(* Logix 5000 project; controller TFF vendor 1 type 14 code 107 rev 34.11; software revision 34.03; part 14 of 36 *)
(* tags used below, declared in another part *)
   ActionCode : DINT;   // Action Code
   ActionValue : REAL;   // Action Value
   Boolean : DINT;   // Boolean Operator
   Branch : BOOL;   // Conditional Branch Flag
   Clear : BOOL;   // Clear Operation Table Flag
   Criteria1BoolValue : BOOL;   // Criteria 1 Discrete Value
   Criteria1Code : DINT;   // Criteria 1 Code
   Criteria1Met : BOOL;   // Criteria 1 Met
   Criteria1Operator : DINT;   // Criteria 1 Operator
   Criteria1RealValue : REAL;   // Criteria 1 Real Value
   Criteria1Type : BOOL;   // Criteria 1 Type 0=Real, 1=Boolean
   Criteria1Value : REAL;   // Criteria 1 Value
   Criteria2BoolValue : BOOL;   // Criteria 2 Discrete Value
   Criteria2Code : DINT;   // Criteria 2 Code
   Criteria2Met : BOOL;   // Criteria 2 Met
   Criteria2Operator : DINT;   // Criteria 2 Operator
   Criteria2RealValue : REAL;   // Criteria 2 Real Value
   Criteria2Type : BOOL;   // Criteria 2 Type 0=Real, 1=Boolean
   Criteria2Value : REAL;   // Criteria 2 Value
   CriteriaMet : BOOL;   // Criteria Met
   DateTime : DINT[7];   // Date and Time
   ErrorCheck : BOOL;   // Error Check Flag
   LastStep : DINT;   // Last Step
   NextStep : DINT;   // Next Step
   PendingStep : DINT;   // Current Step
   PhaseNumber : DINT;   // Phase FOR NEXT Index
   Run : BOOL;   // Operation Run Status
   sColon : STRING4;   // Colon separator String
   sComma : STRING4;   // Comma String
   sDateTime : STRING25;   // Date and Time String
   sPeriod : STRING4;   // Timer separator String
   sTemp : STRING50;   // Temp String
   Structure : DINT;   // Structure code
   sZero : STRING4;   // Zero String
   Tag : DINT;   // Tag value
   Tenths : DINT;   // Thents (Date and Time management)
   ThisStep : DINT;   // This Step (Error management)
   Value : REAL;   // Temp Value
   AlarmControl : AlarmControl;   // Alarm Control
   CCPSystem : CCPSystem;   // CCP System Data
   CPU_Scanning : BOOL;   // System Scanning Flag
   FirstScanComplete : BOOL;   // First Scan Complete Flag
   HoldTime : ALIAS FOR Timers[20];   // Hold Time
   Operation : Operation[6,251];   // Operation Table
   Phase : Phases[6];   // Phase Control Array
   Phase0 : ALIAS FOR Phase[0];   // Phase 0
   Phase0_Totalizer_Feed : ALIAS FOR PhaseTotalizer[0];   // Phase 0 Total Feed
   Phase0_Totalizer_Filtrate : ALIAS FOR PhaseTotalizer[6];   // Phase 0 Total Filtrate
   Phase0_Totalizer_Retentate : ALIAS FOR PhaseTotalizer[12];   // Phase 0 Total Retentate
   PhaseTotalizer : PhaseTotalizer[18];   // Phase Totalizers Array
   PLCFault : FaultRecordType;   // PLC Major Fault Record
   ProcedureTime : ALIAS FOR Timers[19];   // Procedure Time
   Prompt : Prompt[7];   // Prompt Array
   TimerControl : TimerControl;   // Timer Control
   Timers : Timers[22];   // Timer Array
   Totalizer : Totalizers[20];   // Totalizers Array
   YA10 : ALIAS FOR DigitalPoint[59];   // PLC Program Major Fault
(* CCPSystem, continued *)

ROUTINE DateTime   (* structured text *)
// System Date and Time Routine
   (* =======================================================================
   	DateTime : 	This routine returns a string value of date and time in the format "MMDDYYYY,HH:MM:SS.x,".
   				The result is stored in the program tag sDateTime.
   				This string will be used by the BufferEvents and BufferSteps routines for time stamping.
   
   	List of treatments
   		- Get system date and time with GSV instruction
   		- Convert the date and time in DINT format to string format
   
   -----------------------------------------------------------------------------------------------------------------------------------------------------
   	History
   		2019-AUG-13 - ACTEMIUM - B. Roch - Initial version for Candidate Release 3.00.00.00.a
   =========================================================================*)
   
   
   (* Get system date and time with GSV instruction
   =========================================================================*)
   
   (*Get the current date and time from the processor*)
   (*The date and time are stored in an array of 7 values*)
   	GSV (WALLCLOCKTIME, , DateTime, DateTime[0]);
   
   (* Convert the date and time in DINT format to string format
   =========================================================================*)
   (*Month*)
   	DTOS (DateTime[1], sDateTime);
   	(*Add leading zero if value is 1 character*)
   	IF sDateTime.LEN = 1 Then;
   		CONCAT (sZero, sDateTime, sDateTime);
   	END_IF;
   (*Day*)
   	DTOS (DateTime[2], sTemp);
   	(*Add leading zero if value is 1 character*)
   	IF sTemp.LEN = 1 Then;
   		CONCAT (sZero, sTemp, sTemp);
   	END_IF;
   	CONCAT (sDateTime, sTemp, sDateTime);
   (*Year*)
   	DTOS (DateTime[0], sTemp);
   	CONCAT (sDateTime, sTemp, sDateTime);
   	CONCAT (sDateTime, sComma, sDateTime);
   (*Hours*)
   	DTOS (DateTime[3], sTemp);
   	(*Add leading zero if value is 1 character*)
   	IF sTemp.LEN = 1 Then;
   		CONCAT (sZero, sTemp, sTemp);
   	END_IF;
   	CONCAT (sDateTime, sTemp, sDateTime);
   	CONCAT (sDateTime, sColon, sDateTime);
   (*Minutes*)
   	DTOS (DateTime[4], sTemp);
   	(*Add leading zero if value is 1 character*)
   	IF sTemp.LEN = 1 Then;
   		CONCAT (sZero, sTemp, sTemp);
   	END_IF;
   	CONCAT (sDateTime, sTemp, sDateTime);
   	CONCAT (sDateTime, sColon, sDateTime);
   (*Seconds*)
   	DTOS (DateTime[5], sTemp);
   	(*Add leading zero if value is 1 character*)
   	IF sTemp.LEN = 1 Then;
   		CONCAT (sZero, sTemp, sTemp);
   	END_IF;
   	CONCAT (sDateTime, sTemp, sDateTime);
   	CONCAT (sDateTime, sPeriod, sDateTime);
   (*Tenth Seconds*)
   	(*Round the microseconds value to tenths seconds*)
   	Tenths := DateTime[6] / 100000;
   	DTOS (Tenths, sTemp);
   	CONCAT (sDateTime, sTemp, sDateTime);
   	CONCAT (sDateTime, sComma, sDateTime);
   
END_ROUTINE

ROUTINE Error   (* structured text *)
// Step Error Checking
   (* =======================================================================
   	Error : This routine loops through all steps of one phase per processor scan to detect an error
   
   	List of treatments
   		- Initialize
   		- Error check processing
   		- Error found
   		- No error found
   
   -----------------------------------------------------------------------------------------------------------------------------------------------------
   	History
   		2019-AUG-13 - ACTEMIUM - B. Roch - Initial version for Candidate Release 3.00.00.00.a
   		2019-SEP-09 - ACTEMIUM - Q. Spindler - Modifications for Candidate Release 3.00.00.00.c
   					- Change Error check for Criterias and Action Value to -999999.99
   =========================================================================*)
   
   
   (* Initialize
   =========================================================================*)
   (*Initialize error check values first time*)
   IF NOT ErrorCheck THEN;
   	CCPSystem.Error := 0;
   	CCPSystem.ErrorStep:= 0;
   	CCPSystem.ErrorPhase := 0;
   	PhaseNumber := 0;
   	ErrorCheck := 1;
   ELSE;
   	PhaseNumber := PhaseNumber + 1;
   END_IF;
   (* PhaseNumber := 5;*)
   (*Reset the total and last step values*)
   Phase[PhaseNumber].TotalSteps := 0;
   LastStep := 0;
   
   (* Error check processing
   =========================================================================*)
   (*Loop through the steps.  If step number is zero, complete*)
   FOR PendingStep := 1 TO 250 DO;
   	IF Operation[PhaseNumber, PendingStep].Step = 0 THEN;
   		EXIT;
   	END_IF;
   
   	(*Step Number Error Check*)
   	(*Verify step number is equal to or one greater than the previous step number*)
   	ThisStep := Operation[PhaseNumber, PendingStep].Step;
   	IF ThisStep <> LastStep + 1 AND ThisStep <> LastStep THEN;
   		CCPSystem.Error := 1;
   		EXIT;
   	END_IF;
   	LastStep := ThisStep;
   	Phase[PhaseNumber].TotalSteps := PendingStep;
   
   	(*Criteria 1 Error Check*)
   	JSR (Criteria1);
   	IF CCPSystem.Error <> 0 THEN;
   		EXIT;
   	END_IF;
   	IF Criteria1Operator <> 0 AND Criteria1Operator <> 1 AND Criteria1Operator <> 2 AND Criteria1Operator <> 4 THEN;
   		CCPSystem.Error := 3;
   		EXIT;
   	ELSIF Boolean > 2 THEN;
   		CCPSystem.Error := 4;
   		EXIT;
   	ELSIF Criteria1Value = -999999.99 THEN;
   		CCPSystem.Error := 9;
   		EXIT;
   	END_IF;
   
   	(*Criteria 2 Error Check*)
   	JSR (Criteria2);
   	IF CCPSystem.Error <> 0 THEN;
   		EXIT;
   	END_IF;
   	IF Criteria2Operator <> 0 AND Criteria2Operator <> 1 AND Criteria2Operator <> 2 AND Criteria2Operator <> 4 THEN;
   		CCPSystem.Error := 6;
   		EXIT;
   	ELSIF Criteria2Value = -999999.99 THEN;
   		CCPSystem.Error := 10;
   		EXIT;
   	END_IF;
   
   	(*Action Error Check*)
   	JSR (Action);
   	IF CCPSystem.Error <> 0 THEN;
   		EXIT;
   	END_IF;
   	IF ActionValue = -999999.99 THEN;
   		CCPSystem.Error := 11;
   		EXIT;
   	END_IF;
   
   	(*Label Error Check*)
   	IF  Operation[PhaseNumber, PendingStep].Label > 20 THEN;
   		CCPSystem.Error := 8;
   		EXIT;
   	END_IF;
   END_FOR;
   
   (* Error found
   =========================================================================*)
   (*Error Found. Set state to 13, record step and phase number, clear error check flag*)
   IF CCPSystem.Error <> 0 THEN;
   	ErrorCheck := 0;
   	CCPSystem.State := 13;
   	CCPSystem.ErrorStep := PendingStep;
   	CCPSystem.ErrorPhase := PhaseNumber;
   END_IF;
   
   (* No error found
   =========================================================================*)
   (*Complete with no errors. Set state to 0 and clear error check flag*)
   IF PhaseNumber = 5 AND CCPSystem.Error = 0 THEN;
   	ErrorCheck := 0;
   	CCPSystem.State := 0;
   	DTOS (0, CCPSystem.BufferSteps[0]);
   END_IF;
END_ROUTINE

ROUTINE FaultRoutine   (* ladder *)
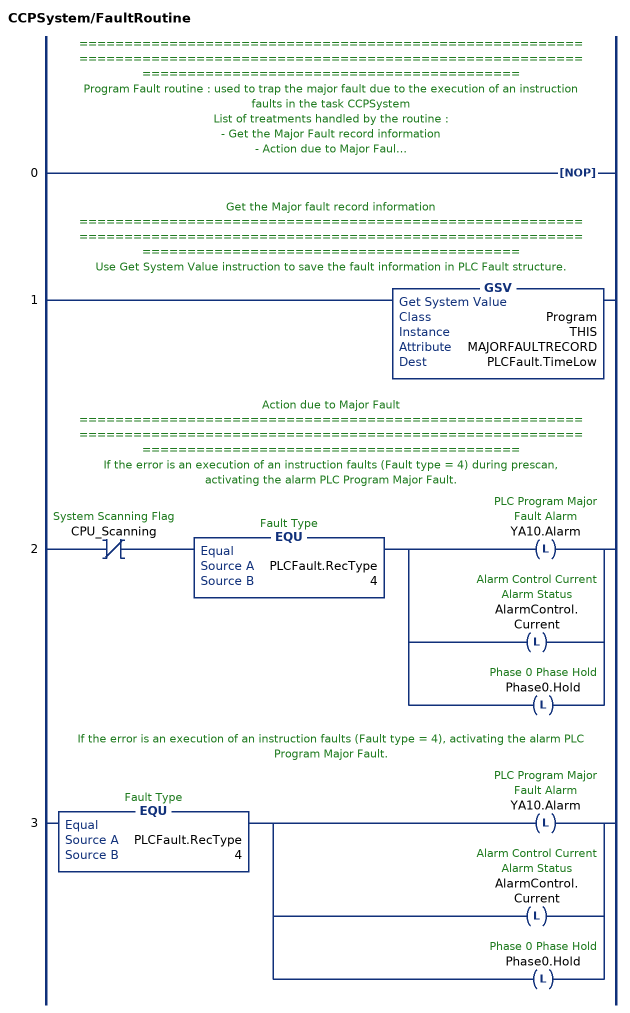
   // ==========================================================================================================================================================
   //                                                            Program Fault routine : used to trap the major fault due to the execution of an instruction faults in the task CCPSystem
   //                                                     List of treatments handled by the routine :
   //                                                          - Get the Major Fault record information
   //                                                          - Action due to Major Fault
   //                                                     -----------------------------------------------------------------------------------------------------------------------------------------------------
   //                                                     History
   //                                                         2019-AUG-13 - Actemium - B. Roch - Initial version for Candidate Release 3.00.00.00.a
   // ==========================================================================================================================================================
   0: NOP();
   // Get the Major fault record information
   // ==========================================================================================================================================================
   // Use Get System Value instruction to save the fault information in PLC Fault structure.
   1: GSV(Program,THIS,MAJORFAULTRECORD,PLCFault.TimeLow);
   // Action due to Major Fault
   // ==========================================================================================================================================================
   // If the error is an execution of an instruction faults (Fault type = 4) during prescan, activating the alarm PLC Program Major Fault.
   2: XIO(CPU_Scanning)EQU(PLCFault.RecType,4)[OTL(YA10.Alarm) ,OTL(AlarmControl.Current) ,OTL(Phase0.Hold) ];
   // If the error is an execution of an instruction faults (Fault type = 4), activating the alarm PLC Program Major Fault.
   3: EQU(PLCFault.RecType,4)[OTL(YA10.Alarm) ,OTL(AlarmControl.Current) ,OTL(Phase0.Hold) ];
END_ROUTINE

ROUTINE MainRoutine   (* ladder *)
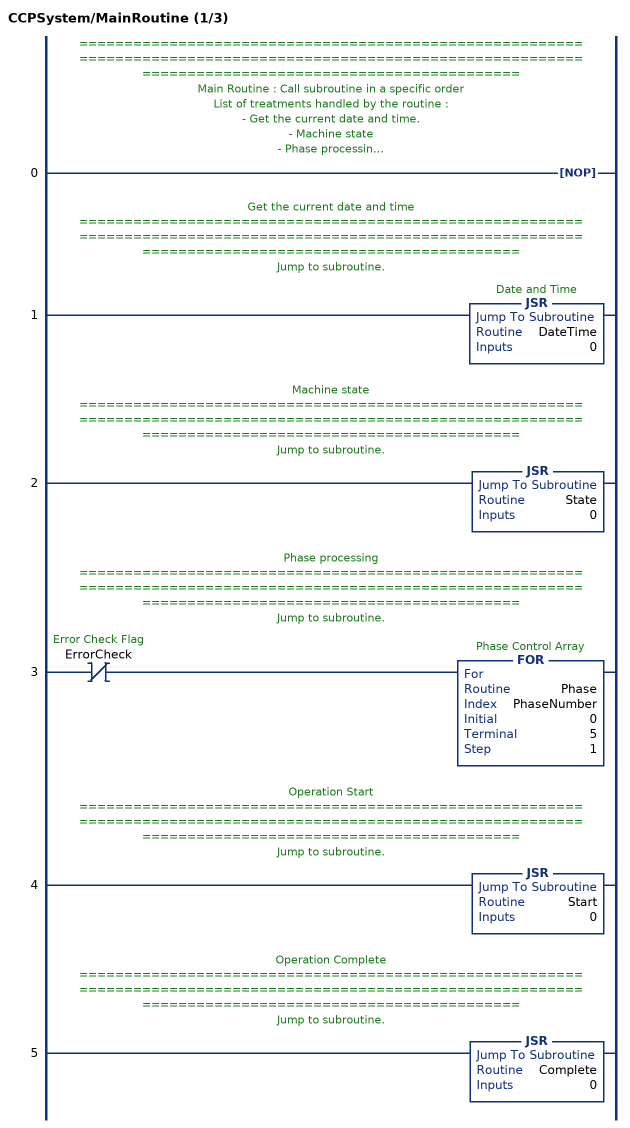
   // ==========================================================================================================================================================
   //                                                                                                            Main Routine : Call subroutine in a specific order
   //                                                     List of treatments handled by the routine :
   //                                                          - Get the current date and time.
   //                                                          - Machine state
   //                                                          - Phase processing
   //                                                          - Operation Start
   //                                                          - Operation Complete
   //                                                          - Procedure timer and totalizer - Hold timer
   //                                                          - Event Log
   //                                                          - CCP System watchdog
   //                                                     -----------------------------------------------------------------------------------------------------------------------------------------------------
   //                                                     History
   //                                                          2019-AUG-13 - Actemium - B. Roch - Initial version for Candidate Release 3.00.00.00.a
   // 2020-SEP-30 - Merck - Q.Spindler - Modifications for Candidate Release 3.00.00.01.a
   // - Add Retentate totalizer
   // ========================================================================================================================================================
   0: NOP();
   // Get the current date and time
   // ==========================================================================================================================================================
   // Jump to subroutine.
   1: JSR(DateTime,0);
   // Machine state
   // ==========================================================================================================================================================
   // Jump to subroutine.
   2: JSR(State,0);
   // Phase processing
   // ==========================================================================================================================================================
   // Jump to subroutine.
   3: XIO(ErrorCheck)FOR(Phase,PhaseNumber,0,5,1);
   // Operation Start
   // ==========================================================================================================================================================
   // Jump to subroutine.
   4: JSR(Start,0);
   // Operation Complete
   // ==========================================================================================================================================================
   // Jump to subroutine.
   5: JSR(Complete,0);
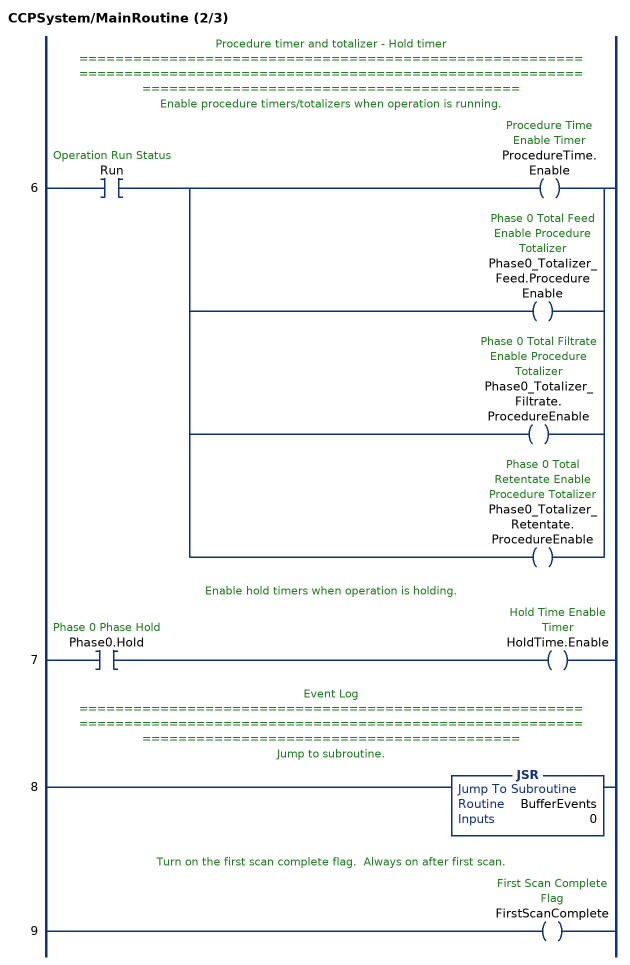
   // Procedure timer and totalizer - Hold timer
   // ==========================================================================================================================================================
   // Enable procedure timers/totalizers when operation is running.
   6: XIC(Run)[OTE(ProcedureTime.Enable) ,OTE(Phase0_Totalizer_Feed.ProcedureEnable) ,OTE(Phase0_Totalizer_Filtrate.ProcedureEnable) ,OTE(Phase0_Totalizer_Retentate.ProcedureEnable) ];
   // Enable hold timers when operation is holding.
   7: XIC(Phase0.Hold)OTE(HoldTime.Enable);
   // Event Log
   // ==========================================================================================================================================================
   // Jump to subroutine.
   8: JSR(BufferEvents,0);
   // Turn on the first scan complete flag.  Always on after first scan.
   9: OTE(FirstScanComplete);
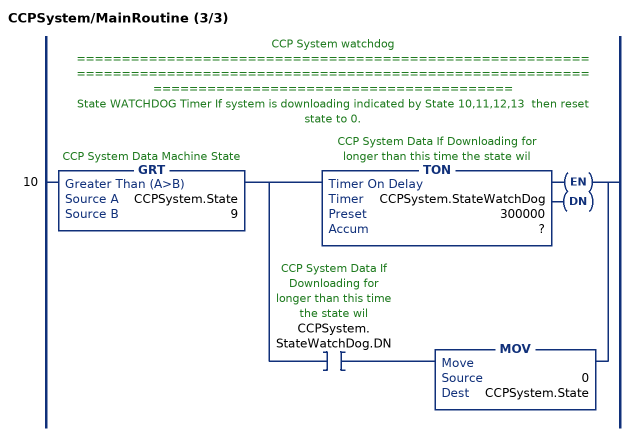
   // CCP System watchdog
   // ==========================================================================================================================================================
   // State WATCHDOG Timer If system is downloading indicated by State 10,11,12,13  then reset state to 0.
   10: GRT(CCPSystem.State,9)[TON(CCPSystem.StateWatchDog,?,?) ,XIC(CCPSystem.StateWatchDog.DN) MOV(0,CCPSystem.State) ];
END_ROUTINE

ROUTINE Phase   (* ladder *)
// Phase Processing Routine
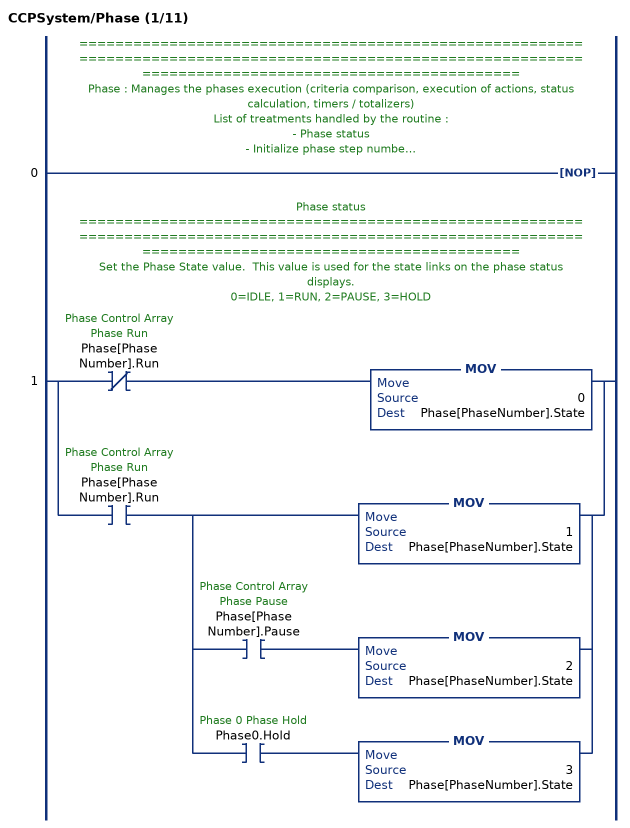
   // ==========================================================================================================================================================
   //                                                                   Phase : Manages the phases execution (criteria comparison, execution of actions, status calculation, timers / totalizers)
   //                                                     List of treatments handled by the routine :
   //                                                          - Phase status
   //                                                          - Initialize phase step number
   //                                                          - Phase Timer / Toalizer
   //                                                          - Phase Stop
   //                                                          - Criteria 1 processing
   //                                                          - Criteria 2 processing
   //                                                          - Jump Step
   //                                                          - Criteria met
   //                                                          - Phase Pause
   //                                                          - Prompt processing
   //                                                          - Branch step processing
   //                                                          - Action processing
   //                                                          - Update step number
   //                                                          - Reset step timer and totalizer
   //                                                     -----------------------------------------------------------------------------------------------------------------------------------------------------
   //                                                     History
   //                                 2019-AUG-13 - Actemium - B. Roch - Initial version for Candidate Release 3.00.00.00.a
   //                                2020-SEP-14 - Merck - Q. Spindler - Modifications for Candidate Release 3.00.00.01.a
   //                                                      - Replace TimerControl.Tick by TimerControl.TickMainTask
   // - Add Retentate totalizer
   // 		               2021-MAY-03 - DAVIDSON- Ch. ARBOGAST - Modifications for Candidate Release 3.01.00.00.a
   //  			- on rung 19 "Reset the step timers...", add "CLR Phase[PhaseNumber].Crit1MetTime"
   //                                          2023-FEB-07 - Davidson - Ch.ARBOGAST - Modifications for Candidate Release 3.02.00.00.a
   //                                                                       - Rung 8. add Hold condition for criteria 1 met Timer (block timer if system in Hold)
   // ========================================================================================================================================================
   0: NOP();
   // Phase status
   // ==========================================================================================================================================================
   // Set the Phase State value.  This value is used for the state links on the phase status displays.
   // 0=IDLE, 1=RUN, 2=PAUSE, 3=HOLD
   1: [XIO(Phase[PhaseNumber].Run) MOV(0,Phase[PhaseNumber].State) ,XIC(Phase[PhaseNumber].Run) [MOV(1,Phase[PhaseNumber].State) ,XIC(Phase[PhaseNumber].Pause) MOV(2,Phase[PhaseNumber].State) ,XIC(Phase0.Hold) MOV(3,Phase[PhaseNumber].State) ] ];
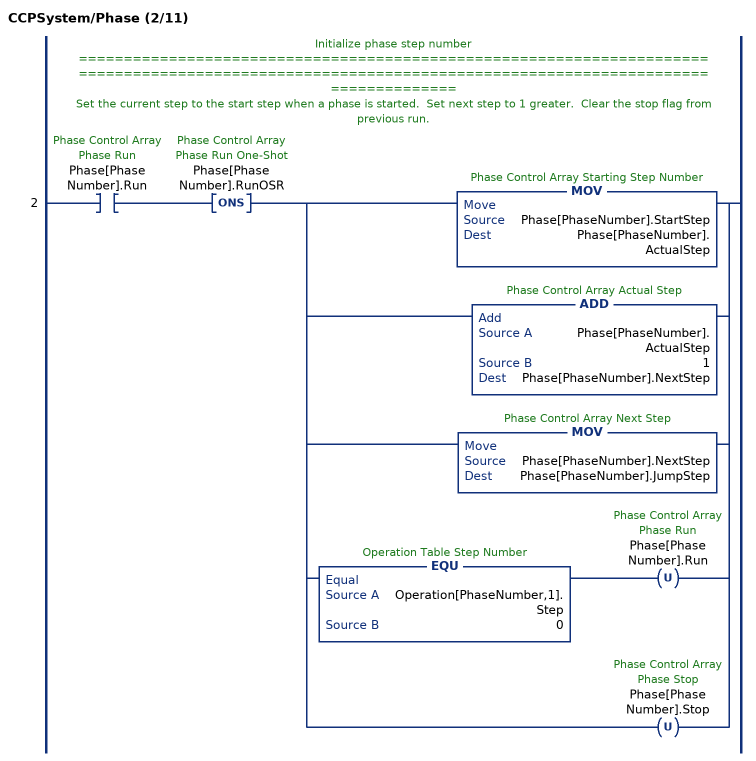
   // Initialize phase step number
   // ==========================================================================================================================================================
   // Set the current step to the start step when a phase is started.  Set next step to 1 greater.  Clear the stop flag from previous run.
   2: XIC(Phase[PhaseNumber].Run)ONS(Phase[PhaseNumber].RunOSR)[MOV(Phase[PhaseNumber].StartStep,Phase[PhaseNumber].ActualStep) ,ADD(Phase[PhaseNumber].ActualStep,1,Phase[PhaseNumber].NextStep) ,MOV(Phase[PhaseNumber].NextStep,Phase[PhaseNumber].JumpStep) ,EQU(Operation[PhaseNumber,1].Step,0) OTU(Phase[PhaseNumber].Run) ,OTU(Phase[PhaseNumber].Stop) ];
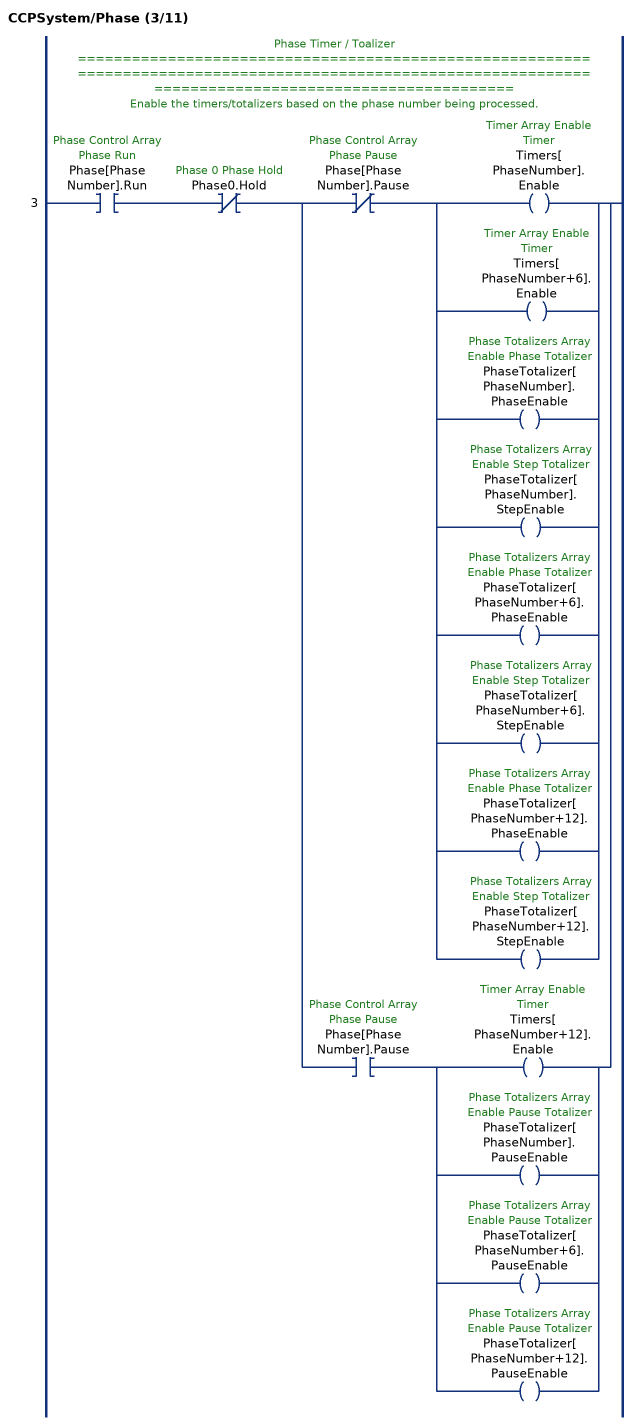
   // Phase Timer / Toalizer
   // ==========================================================================================================================================================
   // Enable the timers/totalizers based on the phase number being processed.
   3: XIC(Phase[PhaseNumber].Run)XIO(Phase0.Hold)[XIO(Phase[PhaseNumber].Pause) [OTE(Timers[PhaseNumber].Enable) ,OTE(Timers[PhaseNumber+6].Enable) ,OTE(PhaseTotalizer[PhaseNumber].PhaseEnable) ,OTE(PhaseTotalizer[PhaseNumber].StepEnable) ,OTE(PhaseTotalizer[PhaseNumber+6].PhaseEnable) ,OTE(PhaseTotalizer[PhaseNumber+6].StepEnable) ,OTE(PhaseTotalizer[PhaseNumber+12].PhaseEnable) ,OTE(PhaseTotalizer[PhaseNumber+12].StepEnable) ] ,XIC(Phase[PhaseNumber].Pause) [OTE(Timers[PhaseNumber+12].Enable) ,OTE(PhaseTotalizer[PhaseNumber].PauseEnable) ,OTE(PhaseTotalizer[PhaseNumber+6].PauseEnable) ,OTE(PhaseTotalizer[PhaseNumber+12].PauseEnable) ] ];
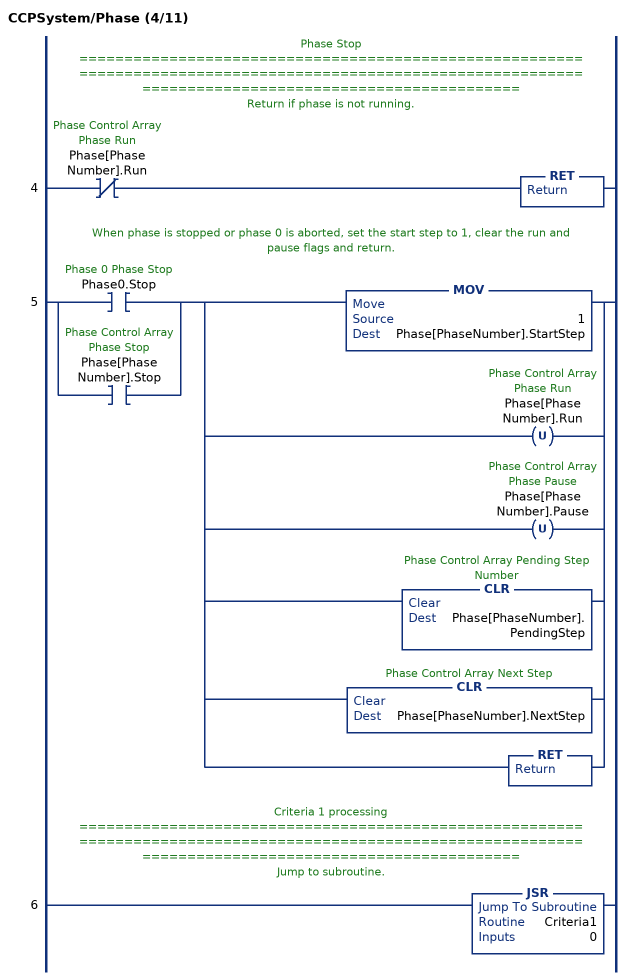
   // Phase Stop
   // ==========================================================================================================================================================
   // Return if phase is not running.
   4: XIO(Phase[PhaseNumber].Run)RET();
   // When phase is stopped or phase 0 is aborted, set the start step to 1, clear the run and pause flags and return.
   5: [XIC(Phase0.Stop) ,XIC(Phase[PhaseNumber].Stop) ][MOV(1,Phase[PhaseNumber].StartStep) ,OTU(Phase[PhaseNumber].Run) ,OTU(Phase[PhaseNumber].Pause) ,CLR(Phase[PhaseNumber].PendingStep) ,CLR(Phase[PhaseNumber].NextStep) ,RET() ];
   // Criteria 1 processing
   // ==========================================================================================================================================================
   // Jump to subroutine.
   6: JSR(Criteria1,0);
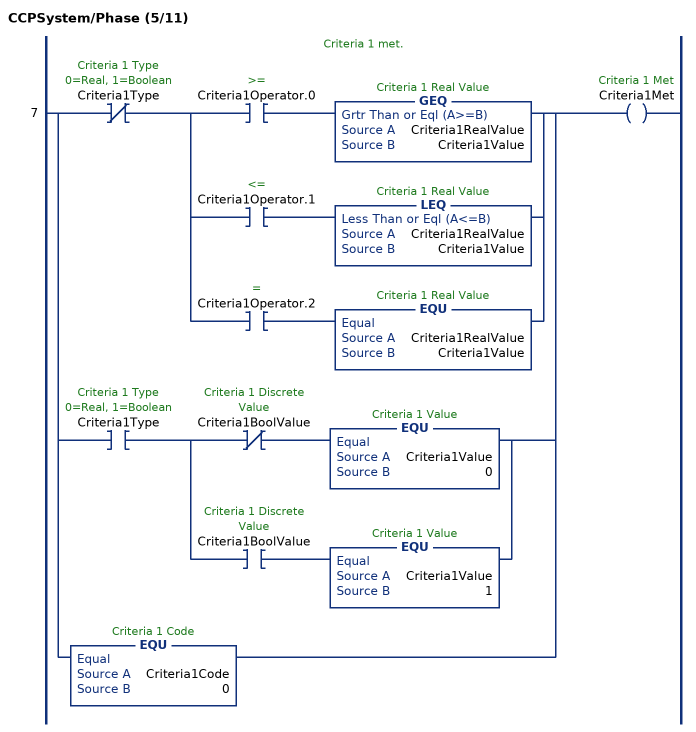
   // Criteria 1 met.
   7: [XIO(Criteria1Type) [XIC(Criteria1Operator.0) GEQ(Criteria1RealValue,Criteria1Value) ,XIC(Criteria1Operator.1) LEQ(Criteria1RealValue,Criteria1Value) ,XIC(Criteria1Operator.2) EQU(Criteria1RealValue,Criteria1Value) ] ,XIC(Criteria1Type) [XIO(Criteria1BoolValue) EQU(Criteria1Value,0) ,XIC(Criteria1BoolValue) EQU(Criteria1Value,1) ] ,EQU(Criteria1Code,0) ]OTE(Criteria1Met);
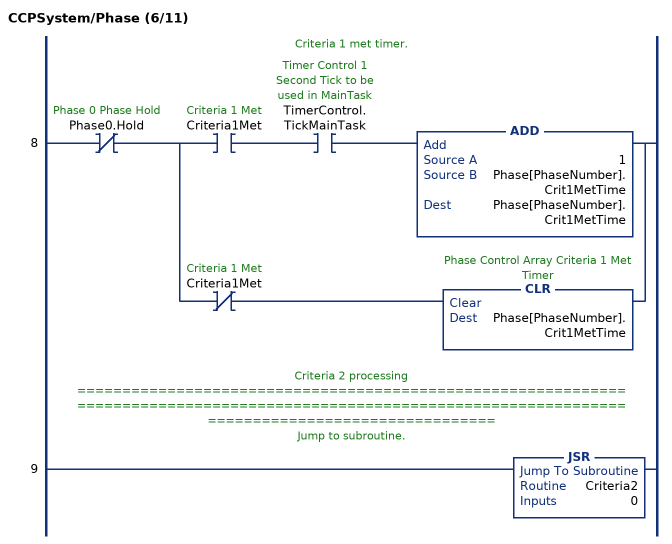
   // Criteria 1 met timer.
   8: XIO(Phase0.Hold)[XIC(Criteria1Met) XIC(TimerControl.TickMainTask) ADD(1,Phase[PhaseNumber].Crit1MetTime,Phase[PhaseNumber].Crit1MetTime) ,XIO(Criteria1Met) CLR(Phase[PhaseNumber].Crit1MetTime) ];
   // Criteria 2 processing
   // ==========================================================================================================================================================
   // Jump to subroutine.
   9: JSR(Criteria2,0);
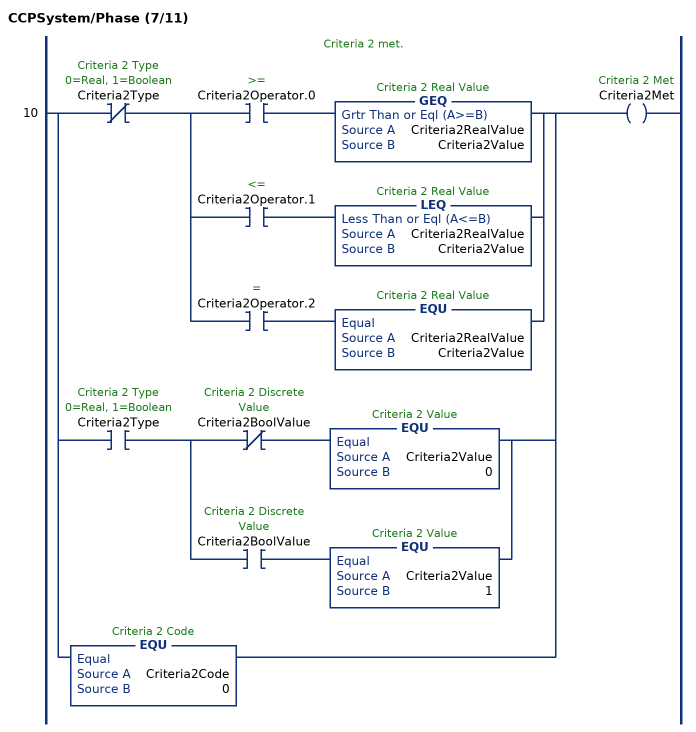
   // Criteria 2 met.
   10: [XIO(Criteria2Type) [XIC(Criteria2Operator.0) GEQ(Criteria2RealValue,Criteria2Value) ,XIC(Criteria2Operator.1) LEQ(Criteria2RealValue,Criteria2Value) ,XIC(Criteria2Operator.2) EQU(Criteria2RealValue,Criteria2Value) ] ,XIC(Criteria2Type) [XIO(Criteria2BoolValue) EQU(Criteria2Value,0) ,XIC(Criteria2BoolValue) EQU(Criteria2Value,1) ] ,EQU(Criteria2Code,0) ]OTE(Criteria2Met);
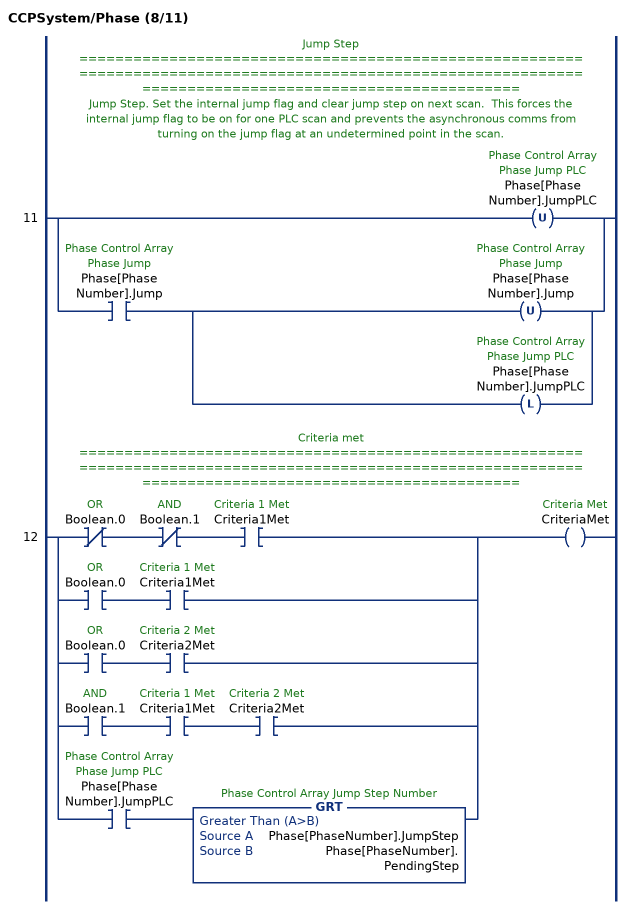
   // Jump Step
   // ==========================================================================================================================================================
   // Jump Step. Set the internal jump flag and clear jump step on next scan.  This forces the internal jump flag to be on for one PLC scan and prevents the asynchronous comms from turning on the jump flag at an undetermined point in the scan.
   11: [OTU(Phase[PhaseNumber].JumpPLC) ,XIC(Phase[PhaseNumber].Jump) [OTU(Phase[PhaseNumber].Jump) ,OTL(Phase[PhaseNumber].JumpPLC) ] ];
   // Criteria met
   // ==========================================================================================================================================================
   12: [XIO(Boolean.0) XIO(Boolean.1) XIC(Criteria1Met) ,XIC(Boolean.0) XIC(Criteria1Met) ,XIC(Boolean.0) XIC(Criteria2Met) ,XIC(Boolean.1) XIC(Criteria1Met) XIC(Criteria2Met) ,XIC(Phase[PhaseNumber].JumpPLC) GRT(Phase[PhaseNumber].JumpStep,Phase[PhaseNumber].PendingStep) ]OTE(CriteriaMet);
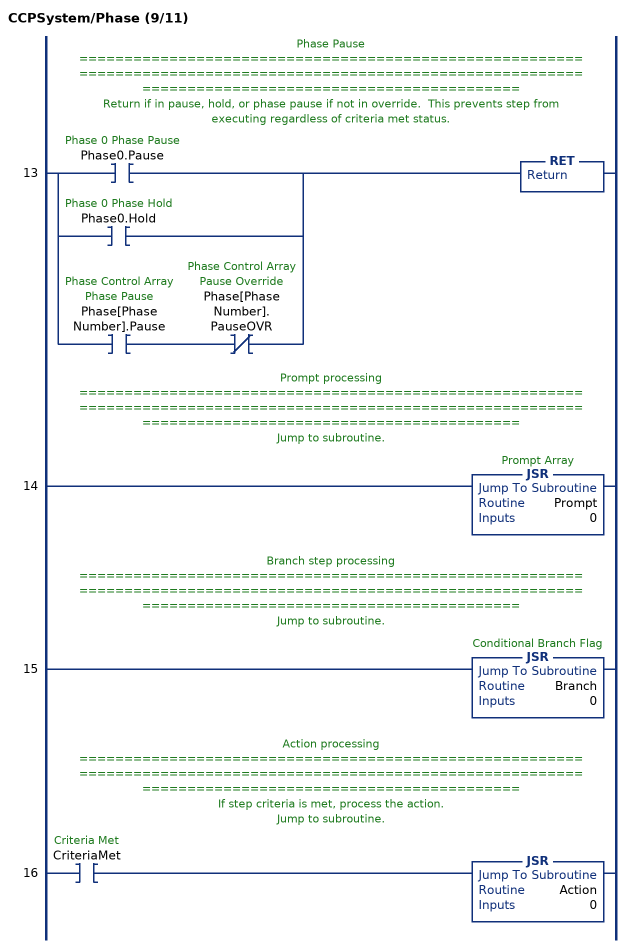
   // Phase Pause
   // ==========================================================================================================================================================
   // Return if in pause, hold, or phase pause if not in override.  This prevents step from executing regardless of criteria met status.
   13: [XIC(Phase0.Pause) ,XIC(Phase0.Hold) ,XIC(Phase[PhaseNumber].Pause) XIO(Phase[PhaseNumber].PauseOVR) ]RET();
   // Prompt processing
   // ==========================================================================================================================================================
   // Jump to subroutine.
   14: JSR(Prompt,0);
   // Branch step processing
   // ==========================================================================================================================================================
   // Jump to subroutine.
   15: JSR(Branch,0);
   // Action processing
   // ==========================================================================================================================================================
   // If step criteria is met, process the action.
   // Jump to subroutine.
   16: XIC(CriteriaMet)JSR(Action,0);
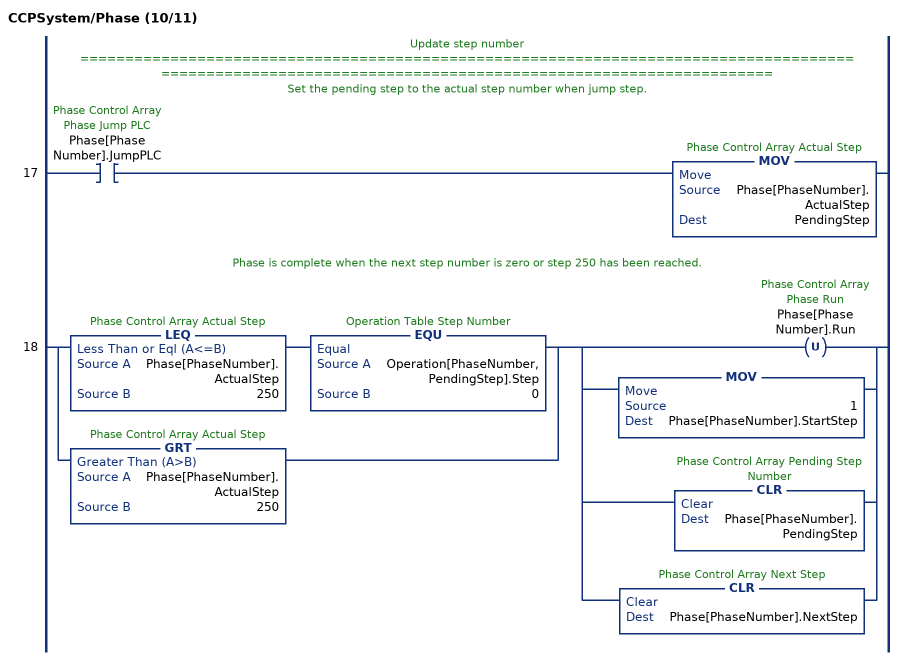
   // Update step number
   // ==========================================================================================================================================================
   // Set the pending step to the actual step number when jump step.
   17: XIC(Phase[PhaseNumber].JumpPLC)MOV(Phase[PhaseNumber].ActualStep,PendingStep);
   // Phase is complete when the next step number is zero or step 250 has been reached.
   18: [LEQ(Phase[PhaseNumber].ActualStep,250) EQU(Operation[PhaseNumber,PendingStep].Step,0) ,GRT(Phase[PhaseNumber].ActualStep,250) ][OTU(Phase[PhaseNumber].Run) ,MOV(1,Phase[PhaseNumber].StartStep) ,CLR(Phase[PhaseNumber].PendingStep) ,CLR(Phase[PhaseNumber].NextStep) ];
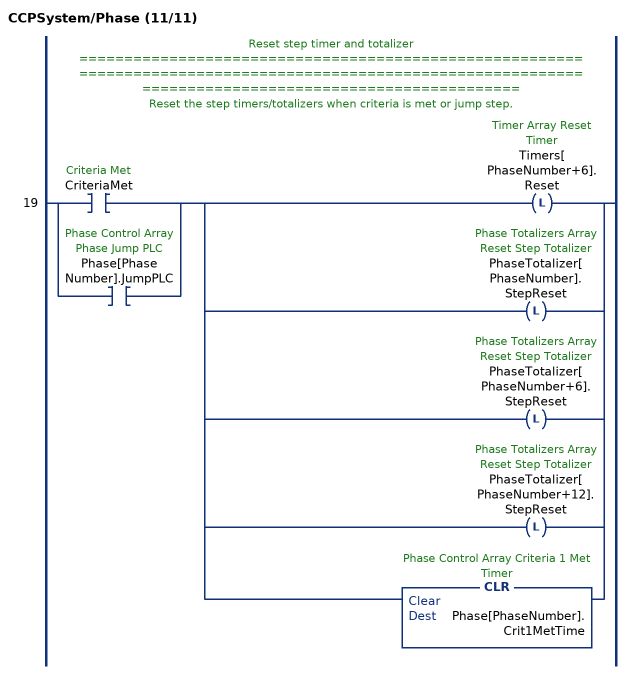
   // Reset step timer and totalizer
   // ==========================================================================================================================================================
   // Reset the step timers/totalizers when criteria is met or jump step.
   19: [XIC(CriteriaMet) ,XIC(Phase[PhaseNumber].JumpPLC) ][OTL(Timers[PhaseNumber+6].Reset) ,OTL(PhaseTotalizer[PhaseNumber].StepReset) ,OTL(PhaseTotalizer[PhaseNumber+6].StepReset) ,OTL(PhaseTotalizer[PhaseNumber+12].StepReset) ,CLR(Phase[PhaseNumber].Crit1MetTime) ];
END_ROUTINE

ROUTINE Prompt   (* ladder *)
// Operator Prompt Routine
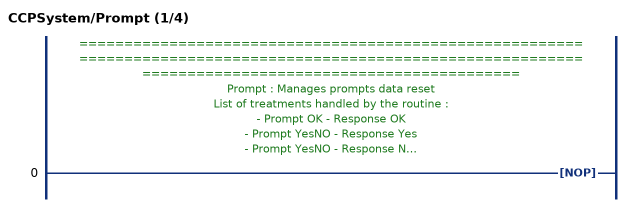
   // ==========================================================================================================================================================
   //                                                                                                                       Prompt : Manages prompts data reset
   //                                                     List of treatments handled by the routine :
   //                                                          - Prompt OK - Response OK
   //                                                          - Prompt YesNO - Response Yes
   //                                                          - Prompt YesNO - Response No
   //                                                     -----------------------------------------------------------------------------------------------------------------------------------------------------
   //                                                     History
   //                                                          2019-AUG-13 - Actemium - B. Roch - Initial version for Candidate Release 3.00.00.00.a
   // 		2023-FEB-08- Davidson - Ch. Arbogast - Modification for Candidate Release 3.02.00.00.a
   //                                            - Rung 1 + 2 + 3:, add condition to avoid discarding the prompt response on other phases than 0
   // ========================================================================================================================================================
   0: NOP();
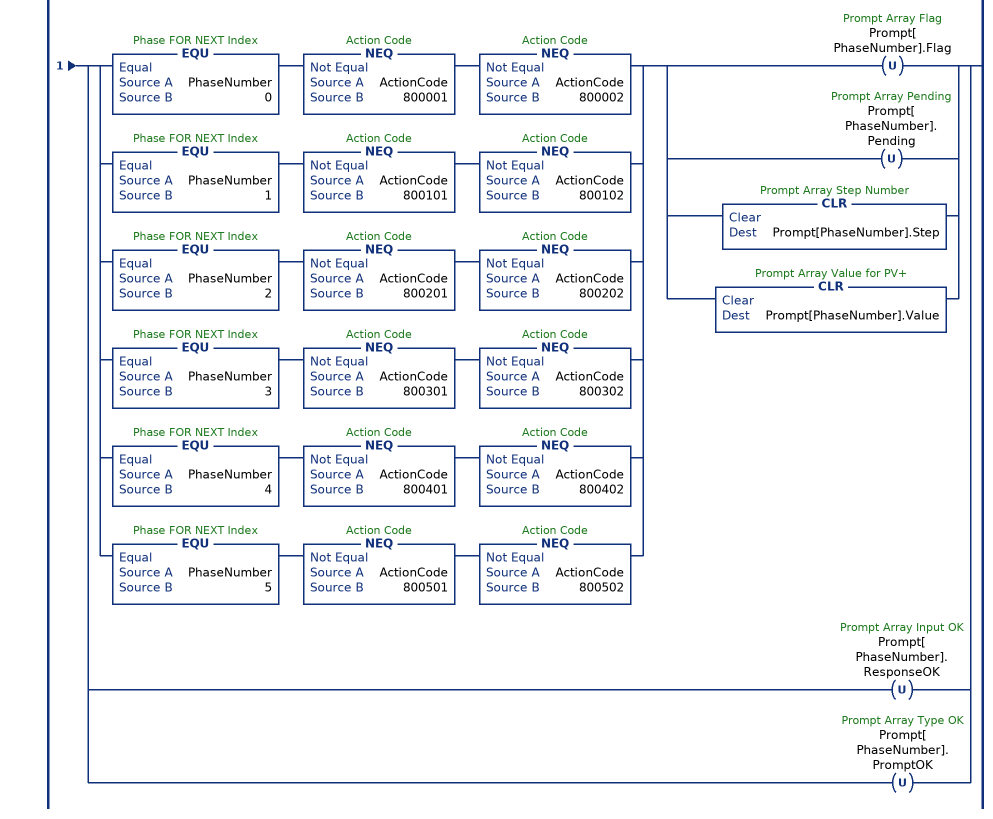
   // Prompt OK - Response OK
   // ==========================================================================================================================================================
   1: XIC(Prompt[PhaseNumber].PromptOK)XIC(Prompt[PhaseNumber].ResponseOK)[XIC(CriteriaMet) ,XIC(Phase[PhaseNumber].JumpPLC) ,EQU(PhaseNumber,0) NEQ(Criteria1Code,800003) NEQ(Criteria2Code,800003) ,EQU(PhaseNumber,1) NEQ(Criteria1Code,800103) NEQ(Criteria2Code,800103) ,EQU(PhaseNumber,2) NEQ(Criteria1Code,800203) NEQ(Criteria2Code,800203) ,EQU(PhaseNumber,3) NEQ(Criteria1Code,800303) NEQ(Criteria2Code,800303) ,EQU(PhaseNumber,4) NEQ(Criteria1Code,800403) NEQ(Criteria2Code,800403) ,EQU(PhaseNumber,5) NEQ(Criteria1Code,800503) NEQ(Criteria2Code,800503) ][[EQU(PhaseNumber,0) NEQ(ActionCode,800001) NEQ(ActionCode,800002) ,EQU(PhaseNumber,1) NEQ(ActionCode,800101) NEQ(ActionCode,800102) ,EQU(PhaseNumber,2) NEQ(ActionCode,800201) NEQ(ActionCode,800202) ,EQU(PhaseNumber,3) NEQ(ActionCode,800301) NEQ(ActionCode,800302) ,EQU(PhaseNumber,4) NEQ(ActionCode,800401) NEQ(ActionCode,800402) ,EQU(PhaseNumber,5) NEQ(ActionCode,800501) NEQ(ActionCode,800502) ] [OTU(Prompt[PhaseNumber].Flag) ,OTU(Prompt[PhaseNumber].Pending) ,CLR(Prompt[PhaseNumber].Step) ,CLR(Prompt[PhaseNumber].Value) ] ,OTU(Prompt[PhaseNumber].ResponseOK) ,OTU(Prompt[PhaseNumber].PromptOK) ];
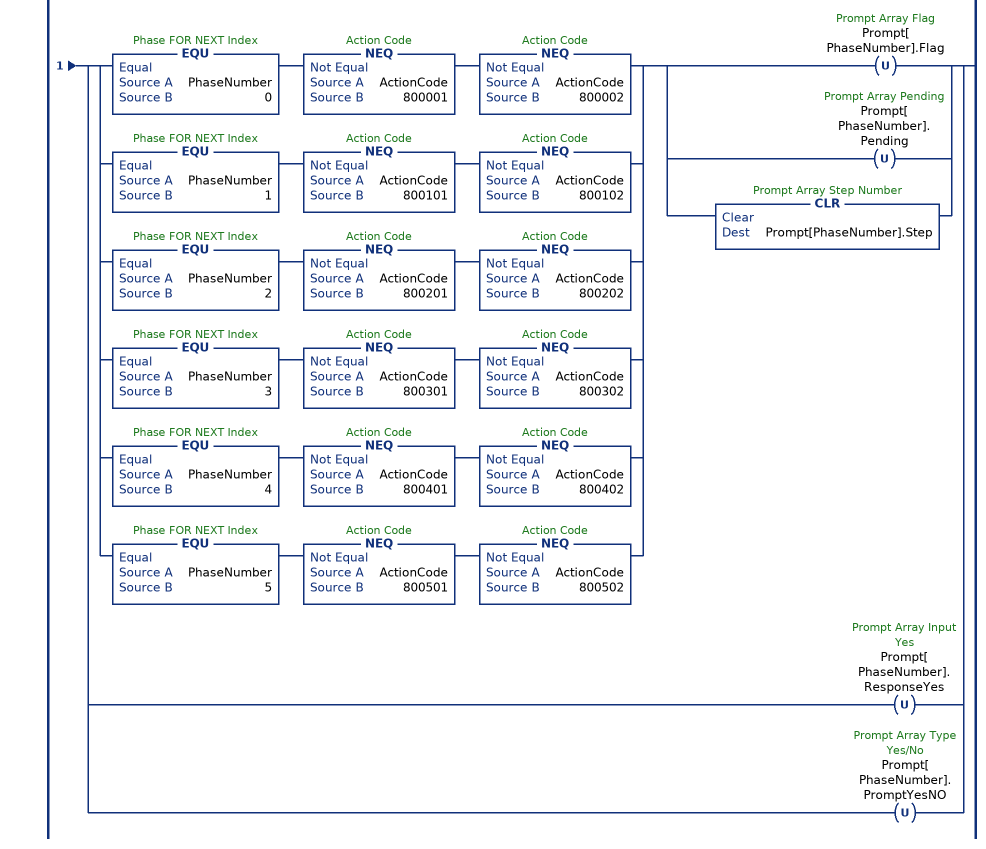
   // Prompt YesNO - Response Yes
   // ==========================================================================================================================================================
   2: XIC(Prompt[PhaseNumber].PromptYesNO)XIC(Prompt[PhaseNumber].ResponseYes)[XIC(CriteriaMet) ,XIC(Phase[PhaseNumber].JumpPLC) ,EQU(PhaseNumber,0) NEQ(Criteria1Code,800004) NEQ(Criteria2Code,800004) ,EQU(PhaseNumber,1) NEQ(Criteria1Code,800104) NEQ(Criteria2Code,800104) ,EQU(PhaseNumber,2) NEQ(Criteria1Code,800204) NEQ(Criteria2Code,800204) ,EQU(PhaseNumber,3) NEQ(Criteria1Code,800304) NEQ(Criteria2Code,800304) ,EQU(PhaseNumber,4) NEQ(Criteria1Code,800404) NEQ(Criteria2Code,800404) ,EQU(PhaseNumber,5) NEQ(Criteria1Code,800504) NEQ(Criteria2Code,800504) ][[EQU(PhaseNumber,0) NEQ(ActionCode,800001) NEQ(ActionCode,800002) ,EQU(PhaseNumber,1) NEQ(ActionCode,800101) NEQ(ActionCode,800102) ,EQU(PhaseNumber,2) NEQ(ActionCode,800201) NEQ(ActionCode,800202) ,EQU(PhaseNumber,3) NEQ(ActionCode,800301) NEQ(ActionCode,800302) ,EQU(PhaseNumber,4) NEQ(ActionCode,800401) NEQ(ActionCode,800402) ,EQU(PhaseNumber,5) NEQ(ActionCode,800501) NEQ(ActionCode,800502) ] [OTU(Prompt[PhaseNumber].Flag) ,OTU(Prompt[PhaseNumber].Pending) ,CLR(Prompt[PhaseNumber].Step) ] ,OTU(Prompt[PhaseNumber].ResponseYes) ,OTU(Prompt[PhaseNumber].PromptYesNO) ];
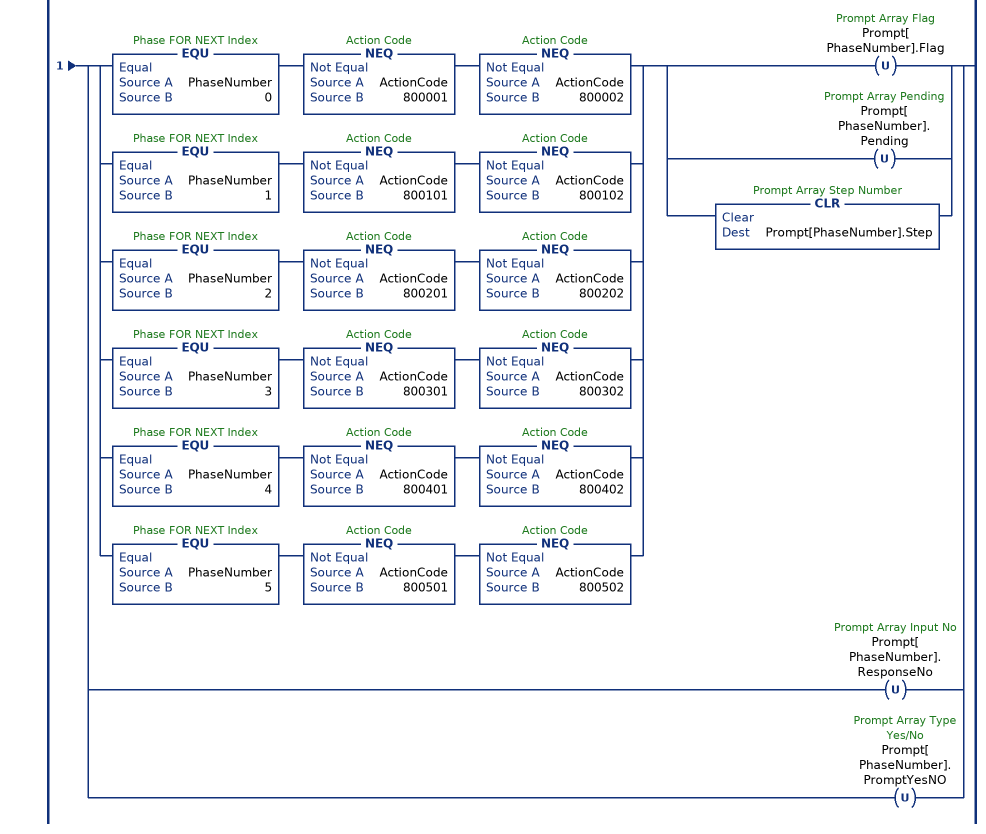
   // Prompt YesNO - Response No
   // ==========================================================================================================================================================
   3: XIC(Prompt[PhaseNumber].PromptYesNO)XIC(Prompt[PhaseNumber].ResponseNo)[XIC(CriteriaMet) ,XIC(Phase[PhaseNumber].JumpPLC) ,EQU(PhaseNumber,0) NEQ(Criteria1Code,800005) NEQ(Criteria2Code,800005) ,EQU(PhaseNumber,1) NEQ(Criteria1Code,800105) NEQ(Criteria2Code,800105) ,EQU(PhaseNumber,2) NEQ(Criteria1Code,800205) NEQ(Criteria2Code,800205) ,EQU(PhaseNumber,3) NEQ(Criteria1Code,800305) NEQ(Criteria2Code,800305) ,EQU(PhaseNumber,4) NEQ(Criteria1Code,800405) NEQ(Criteria2Code,800405) ,EQU(PhaseNumber,5) NEQ(Criteria1Code,800505) NEQ(Criteria2Code,800505) ][[EQU(PhaseNumber,0) NEQ(ActionCode,800001) NEQ(ActionCode,800002) ,EQU(PhaseNumber,1) NEQ(ActionCode,800101) NEQ(ActionCode,800102) ,EQU(PhaseNumber,2) NEQ(ActionCode,800201) NEQ(ActionCode,800202) ,EQU(PhaseNumber,3) NEQ(ActionCode,800301) NEQ(ActionCode,800302) ,EQU(PhaseNumber,4) NEQ(ActionCode,800401) NEQ(ActionCode,800402) ,EQU(PhaseNumber,5) NEQ(ActionCode,800501) NEQ(ActionCode,800502) ] [OTU(Prompt[PhaseNumber].Flag) ,OTU(Prompt[PhaseNumber].Pending) ,CLR(Prompt[PhaseNumber].Step) ] ,OTU(Prompt[PhaseNumber].ResponseNo) ,OTU(Prompt[PhaseNumber].PromptYesNO) ];
END_ROUTINE
